{region 'Documentation'}
(*!
<summary>Composes two minimal real Test Cases with the real production Orchestrator.</summary>
<description>
Only publisher binding and call counters are added for observation.
The inherited base and real helper own all transitions, requests and reservations.
Children are initialized once in Configure, then Reset and executed twice without rebinding.
</description>
*)
{endregion}
FUNCTION_BLOCK SuiteIntegrationSubject EXTENDS TestSuiteBase
VAR
    FFirst : SuiteIntegrationChild;
    FSecond : SuiteIntegrationChild;
    FTestCases : ARRAY[4..6] OF I_TestCase;
    FRealOrchestrator : OrchestratorProbe;
    FBodyCallCount : UDINT;
    FConfigureCount : UINT;
END_VAR

FBodyCallCount := FBodyCallCount + 1;
SUPER^();

{region 'Documentation'}
(*!
<summary>Binds every producer before Initialize; never modifies the global publisher.</summary>
*)
{endregion}
METHOD PUBLIC BindPublisher
VAR_INPUT
    Publisher : I_EventPublisher; //! Nonzero isolated event publisher retained before subject initialization; keep it alive through all subject use.
END_VAR
FEventPublisher := Publisher;
FRealOrchestrator.BindPublisher(Publisher := Publisher);
FOrchestrator := FRealOrchestrator;
FFirst.BindPublisher(Publisher := Publisher);
FSecond.BindPublisher(Publisher := Publisher);
FBodyCallCount := 0;
FConfigureCount := 0;
END_METHOD

{region 'Documentation'}
(*!
<summary>Confirms one concrete child call per Suite call, including Reset and Completed.</summary>
*)
{endregion}
{attribute 'monitoring' := 'call'}
PROPERTY PUBLIC ChildCallsMatch : BOOL //! Confirms one concrete child call per Suite call, including Reset and Completed.
GET
ChildCallsMatch := (FFirst.BodyCallCount = FBodyCallCount) AND (FSecond.BodyCallCount = FBodyCallCount);
END_GET
END_PROPERTY

{region 'Documentation'}
(*!
<summary>Initializes and registers two real children serially in a shifted array with one unused slot.</summary>
*)
{endregion}
METHOD PROTECTED Configure
VAR_IN_OUT
    // SA0167: Borrowed setup builder; no temporary instance is created.
    {attribute 'analysis' := '-167'}
    Builder : TestSuiteConfigurationBuilder; //! Borrowed owner configuration builder used only during this Configure call; register this owner's concrete children.
END_VAR
VAR
    Config : ST_TestCaseConfig;
END_VAR
FConfigureCount := FConfigureCount + 1;
Builder.Initialize(Mode := E_OrchestrationMode.Serial,
    TestCases := FTestCases);
FFirst.Initialize(Parent := THIS^,
    TestName := 'First',
    Config := Config);
FSecond.Initialize(Parent := THIS^,
    TestName := 'Second',
    Config := Config);
Builder.Register(TestCase := FFirst);
Builder.Register(TestCase := FSecond);
END_METHOD

{region 'Documentation'}
(*!
<summary>Distinguishes Reset/repeat from reinitializing the subject.</summary>
*)
{endregion}
{attribute 'monitoring' := 'call'}
PROPERTY PUBLIC ConfigureCount : UINT //! Distinguishes Reset/repeat from reinitializing the subject.
GET
ConfigureCount := FConfigureCount;
END_GET
END_PROPERTY

{region 'Documentation'}
(*!
<summary>Resolves the actual registered array index without executing the child.</summary>
*)
{endregion}
METHOD PUBLIC GetTestCase : I_TestCase //! Typed child interface at the original array index; zero when no entry is available.
VAR_INPUT
    Index : DINT; //! Original occupied child-array index, rather than an ordinal position.
END_VAR
GetTestCase := 0;
IF (ChildCount = 0) OR (Index < ChildArrayLowerBound)
    OR (DINT_TO_LINT(Index) >= DINT_TO_LINT(ChildArrayLowerBound) + UINT_TO_LINT(ChildCount)) THEN
    RETURN;
END_IF;
GetTestCase := FTestCases[Index];
END_METHOD

{region 'Documentation'}
(*!
<summary>Calls both children once per initialized Suite call; the helper requests their lifecycle actions.</summary>
*)
{endregion}
METHOD PROTECTED ProcessTestCases
FFirst();
FSecond();
END_METHOD

END_FUNCTION_BLOCK

(* stored: Version 1.1.0.1
   POU SuiteIntegrationSubject: Id {279ede58-4fe0-45a2-9b27-f0adb5bf63f3}, SpecialFunc None
   Folder Internal: Id {243039e3-c84c-4097-a8ac-7891f5cce17d}
   Method BindPublisher: Id {2f7a0930-a534-4e96-8378-6ea9b9244232}
   Property ChildCallsMatch: Id {a592d272-097e-49cc-beb5-8e240156365b}
   Get Get: Id {d76d69a8-d1b9-40a6-a4b2-9923af3586f0}
   Method Configure: Id {67e63565-4a71-4020-bf96-df1e458c6834}
   Property ConfigureCount: Id {a8e76c12-e820-4095-b5fc-8ab931be9474}
   Get Get: Id {90f8a366-d48f-4b53-a7ad-dfc5daed9980}
   Method GetTestCase: Id {1aa83588-01a5-49b3-898e-16781b00462b}
   Method ProcessTestCases: Id {b36c0e43-2b13-41f3-a1db-c84c6f95ea40} *)
